(* IEC 61131-3 sources: kns-port-domestic/tools/port_metrics_tests/fixtures/app/src/POUs/PRG_Main, 1 file *)

(* ---- PRG_Main.decl.st ---- *)
PROGRAM PRG_Main
VAR
    fbPump : FB_Pump;
    xStartCmd : BOOL;
END_VAR
